(* IEC 61131-3 sources: SRCI_CLIENT_PLC/RobotLibrary/Library/POUs/Calculation/MC_CalculateFrame/Structures, 4 files *)

(* ---- CalculateFrameOutCmd.st ---- *)
{attribute 'pack_mode' := '1'}
// -------------------------------------------------------------------------
//  SRCI Robot Library
// -------------------------------------------------------------------------
//
//  Object:      CalculateFrameOutCmd
//  Author:      Thorsten Brach
//  Date:        2024-06-09
//
//  Description:
//
//
//  Copyright:
//    (C) 2024 Thorsten Brach. All rights reserved
//             Licensed under the MIT License.
//
//  Disclaimer:
//    This project is provided without any guarantee and can be used for
//    private and commercial purposes. Any use is at the user’s
//    own risk and responsibility.
//
// -------------------------------------------------------------------------
TYPE CalculateFrameOutCmd :
STRUCT
  /// Date
  IEC_Date       : IEC_DATE;
  /// Time
  IEC_TIME       : IEC_TIME;
  /// Index of frame on which the calculated frame is depending
  /// •      0: WCS (default)
  /// • 1..254: User frames
  ReferenceFrame : USINT;
  /// Position
  Position       : RobotCartesianPositionBase;
END_STRUCT
END_TYPE

(* ---- CalculateFrameParCmd.st ---- *)
{attribute 'pack_mode' := '1'}
// -------------------------------------------------------------------------
//  SRCI Robot Library
// -------------------------------------------------------------------------
//
//  Object:      CalculateFrameParCmd
//  Author:      Thorsten Brach
//  Date:        2024-06-09
//
//  Description:
//
//
//  Copyright:
//    (C) 2024 Thorsten Brach. All rights reserved
//             Licensed under the MIT License.
//
//  Disclaimer:
//    This project is provided without any guarantee and can be used for
//    private and commercial purposes. Any use is at the user’s
//    own risk and responsibility.
//
// -------------------------------------------------------------------------
TYPE CalculateFrameParCmd :
STRUCT
  /// Define which method should be used to calculate the tool frame
  Mode               : FrameCalculationMode;
  /// Index of target frame
  /// • 0: WCS (default)
  /// • 1..254: User frames
  FrameNo            : USINT;
  /// Cartesian position in the positive direction of the  X-Axis of the calculated frame coordinate system relative to the given frame
  Position_X         : RobotCartesianPosition;
  /// Cartesian position in the XY-plane of the calculated frame coordinate system relative to the given frame.
  Position_XY        : RobotCartesianPosition;
  /// Cartesian position of the origin of the calculated frame coordinate system relative to the given frame.
  Origin             : RobotCartesianPosition;
  /// Cartesian position of the postponement of the origin of the calculated frame coordinate system relative to the given frame.
  /// Auxiliary position if the origin of the can’t be reached by the robot, i.e. because it is inside an object.
  OriginShift        : RobotCartesianPosition;
  /// Index of frame on which the calculated frame is depending
  /// •      0: WCS (default)
  /// • 1..254: User frames
  ReferenceFrame     : USINT;
END_STRUCT
END_TYPE

(* ---- CalculateFrameRecvData.st ---- *)
{attribute 'pack_mode' := '1'}
// -------------------------------------------------------------------------
//  SRCI Robot Library
// -------------------------------------------------------------------------
//
//  Object:      CalculateFrameRecvData
//  Author:      Thorsten Brach
//  Date:        2024-06-09
//
//  Description:
//
//
//  Copyright:
//    (C) 2024 Thorsten Brach. All rights reserved
//             Licensed under the MIT License.
//
//  Disclaimer:
//    This project is provided without any guarantee and can be used for
//    private and commercial purposes. Any use is at the user’s
//    own risk and responsibility.
//
// -------------------------------------------------------------------------
TYPE CalculateFrameRecvData EXTENDS RspHeader :
STRUCT
  /// Date
  IEC_Date       : IEC_DATE;
  /// Time
  IEC_TIME       : IEC_TIME;
  /// Index of frame on which the calculated frame is depending
  /// •      0: WCS (default)
  /// • 1..254: User frames
  ReferenceFrame : USINT;
  /// Reserve
  Reserve        : BYTE;
  /// Position
  Position       : RobotCartesianPositionBase;
END_STRUCT
END_TYPE

(* ---- CalculateFrameSendData.st ---- *)
{attribute 'pack_mode' := '1'}
// -------------------------------------------------------------------------
//  SRCI Robot Library
// -------------------------------------------------------------------------
//
//  Object:      CalculateFrameSendData
//  Author:      Thorsten Brach
//  Date:        2024-06-09
//
//  Description:
//
//
//  Copyright:
//    (C) 2024 Thorsten Brach. All rights reserved
//             Licensed under the MIT License.
//
//  Disclaimer:
//    This project is provided without any guarantee and can be used for
//    private and commercial purposes. Any use is at the user’s
//    own risk and responsibility.
//
// -------------------------------------------------------------------------
TYPE CalculateFrameSendData EXTENDS CmdHeader:
STRUCT
  /// Incremented with each position of the input parameter "PositionsArray" sent from the PLC to the RC.
  /// Default: 0
  DataIndex          : USINT;

  /// Set TRUE by the client, when according to the user selected "Mode" the final position of the input parameter "PositionsArray" is sent to the RC.
  /// Default: FALSE
  DataComplete       : BYTE;
  ///
  Reserve            : BYTE;
  /// Index of target frame
  /// • 0: WCS (default)
  /// • 1..254: User frames
  FrameNo            : USINT;
  /// Index of frame on which the calculated frame is depending
  /// •      0: WCS (default)
  /// • 1..254: User frames
  ReferenceFrame     : USINT;
  /// Define which method should be used to calculate the frame coordinate system: M
  /// • 0: Three-Point-Method (default) O
  /// • 1: Four-Point-Method O
  /// • 2: One-Point-Method
  Mode               : SINT;
  /// Cartesian position
  Position           : RobotCartesianPosition;
END_STRUCT
END_TYPE
